(* IEC 61131-3 sources: rusty/tests/lit/ir_tests/include, 1 file *)

(* ---- included_types.st ---- *)
TYPE
    IncludedStruct : STRUCT
        v : DINT;
    END_STRUCT
END_TYPE
